(* IEC 61131-3 sources: trust-platform/examples/OSCAT/weather_station_conversion/non-oop/src, 1 file *)

(* ---- Configuration.st ---- *)
CONFIGURATION WeatherStationConversionClassicConfiguration
RESOURCE WeatherStationConversionClassic ON PLC
    TASK MainTask (INTERVAL := T#1s, PRIORITY := 1);
    PROGRAM Main WITH MainTask : Main;
END_RESOURCE
END_CONFIGURATION
